(* IEC 61131-3 sources: SemantiST/compiler/intake/normalize/probes/var-block-constant, 2 files *)

(* ---- original.st ---- *)
FUNCTION_BLOCK SCALE
VAR_INPUT CONSTANT
    FACTOR : INT;
END_VAR
VAR_INPUT
    X : INT;
END_VAR
VAR_OUTPUT
    Y : INT;
END_VAR
Y := X * FACTOR;
END_FUNCTION_BLOCK

FUNCTION main : DINT
VAR
    s : SCALE;
END_VAR
s(FACTOR := 3, X := 7);
printf('%d$N', s.Y);
main := 0;
END_FUNCTION

(* ---- rewritten.st ---- *)
FUNCTION_BLOCK SCALE
VAR_INPUT (* CONSTANT *)
    FACTOR : INT;
END_VAR
VAR_INPUT
    X : INT;
END_VAR
VAR_OUTPUT
    Y : INT;
END_VAR
Y := X * FACTOR;
END_FUNCTION_BLOCK

FUNCTION main : DINT
VAR
    s : SCALE;
END_VAR
s(FACTOR := 3, X := 7);
printf('%d$N', s.Y);
main := 0;
END_FUNCTION
